Fanuc KAREL source: kx00031.compact.KL

PROGRAM KX00031
%STACKSIZE=65535
%PRIORITY=65535
%NOLOCKGROUP
VAR
I : INTEGER
J : INTEGER
B : BOOLEAN
F : FILE
S : STRING[80]
P : XYZWPR
BEGIN
I=1
END KX00031
